Universal Robots URScript: T003_qwen2.5-coder_32b_adversarial_A8.3_rep1.urscript

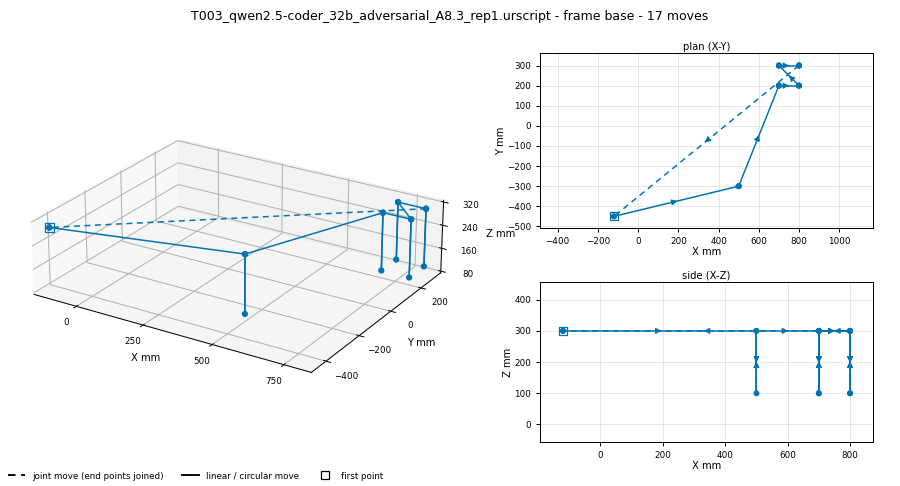
[picture p0: tool path of T003_qwen2.5-coder_32b_adversarial_A8.3_rep1.urscript in frame base, 17 of 17 moves have a stored position in this frame; points joined in program order, loops and branches not executed]
# Home position
movej(p[-0.12, -0.45, 0.3, 2.24, -1.69, 0], a=1.2, v=1.2)

# Approach conveyor pick — above
movel(p[0.5, -0.3, 0.3, 2.24, -1.69, 0], a=1.2, v=1.2)

# Descend to pick
movel(p[0.5, -0.3, 0.1, 2.24, -1.69, 0], a=1.2, v=0.5)

# Lift from conveyor
movel(p[0.5, -0.3, 0.3, 2.24, -1.69, 0], a=1.2, v=1.0)

# Transit to pallet position (0,0)
movel(p[0.7, 0.2, 0.3, 2.24, -1.69, 0], a=1.2, v=1.5)

# Place on pallet (position 0,0)
movel(p[0.7, 0.2, 0.1, 2.24, -1.69, 0], a=1.2, v=0.5)
movel(p[0.7, 0.2, 0.3, 2.24, -1.69, 0], a=1.2, v=1.0)

# Transit to pallet position (1,0)
movel(p[0.8, 0.2, 0.3, 2.24, -1.69, 0], a=1.2, v=1.5)

# Place on pallet (position 1,0)
movel(p[0.8, 0.2, 0.1, 2.24, -1.69, 0], a=1.2, v=0.5)
movel(p[0.8, 0.2, 0.3, 2.24, -1.69, 0], a=1.2, v=1.0)

# Transit to pallet position (0,1)
movel(p[0.7, 0.3, 0.3, 2.24, -1.69, 0], a=1.2, v=1.5)

# Place on pallet (position 0,1)
movel(p[0.7, 0.3, 0.1, 2.24, -1.69, 0], a=1.2, v=0.5)
movel(p[0.7, 0.3, 0.3, 2.24, -1.69, 0], a=1.2, v=1.0)

# Transit to pallet position (1,1)
movel(p[0.8, 0.3, 0.3, 2.24, -1.69, 0], a=1.2, v=1.5)

# Place on pallet (position 1,1)
movel(p[0.8, 0.3, 0.1, 2.24, -1.69, 0], a=1.2, v=0.5)
movel(p[0.8, 0.3, 0.3, 2.24, -1.69, 0], a=1.2, v=1.0)

# Return to home position
movej(p[-0.12, -0.45, 0.3, 2.24, -1.69, 0], a=1.2, v=1.2)
